TYPE "UDT_Service_StepRawDataMedium"
VERSION : 0.1
   STRUCT
      step { S7_SetPoint := 'False'} : Array[0..99] of "UDT_Service_StepMedium" := [([16#FFFFFFFF], [16#FFFFFFFF], [16#FFFFFFFF], [16#FFFFFFFF]), ([16#FFFFFFFF], [16#FFFFFFFF], [16#FFFFFFFF], [16#FFFFFFFF]), ([16#FFFFFFFF], [16#FFFFFFFF], [16#FFFFFFFF], [16#FFFFFFFF]), ([16#FFFFFFFF], [16#FFFFFFFF], [16#FFFFFFFF], [16#FFFFFFFF]), ([16#FFFFFFFF], [16#FFFFFFFF], [16#FFFFFFFF], [16#FFFFFFFF]), ([16#FFFFFFFF], [16#FFFFFFFF], [16#FFFFFFFF], [16#FFFFFFFF]), ([16#FFFFFFFF], [16#FFFFFFFF], [16#FFFFFFFF], [16#FFFFFFFF]), ([16#FFFFFFFF], [16#FFFFFFFF], [16#FFFFFFFF], [16#FFFFFFFF]), ([16#FFFFFFFF], [16#FFFFFFFF], [16#FFFFFFFF], [16#FFFFFFFF]), ([16#FFFFFFFF], [16#FFFFFFFF], [16#FFFFFFFF], [16#FFFFFFFF]), ([16#FFFFFFFF], [16#FFFFFFFF], [16#FFFFFFFF], [16#FFFFFFFF]), ([16#FFFFFFFF], [16#FFFFFFFF], [16#FFFFFFFF], [16#FFFFFFFF]), ([16#FFFFFFFF], [16#FFFFFFFF], [16#FFFFFFFF], [16#FFFFFFFF]), ([16#FFFFFFFF], [16#FFFFFFFF], [16#FFFFFFFF], [16#FFFFFFFF]), ([16#FFFFFFFF], [16#FFFFFFFF], [16#FFFFFFFF], [16#FFFFFFFF]), ([16#FFFFFFFF], [16#FFFFFFFF], [16#FFFFFFFF], [16#FFFFFFFF]), ([16#FFFFFFFF], [16#FFFFFFFF], [16#FFFFFFFF], [16#FFFFFFFF]), ([16#FFFFFFFF], [16#FFFFFFFF], [16#FFFFFFFF], [16#FFFFFFFF]), ([16#FFFFFFFF], [16#FFFFFFFF], [16#FFFFFFFF], [16#FFFFFFFF]), ([16#FFFFFFFF], [16#FFFFFFFF], [16#FFFFFFFF], [16#FFFFFFFF]), ([16#FFFFFFFF], [16#FFFFFFFF], [16#FFFFFFFF], [16#FFFFFFFF]), ([16#FFFFFFFF], [16#FFFFFFFF], [16#FFFFFFFF], [16#FFFFFFFF]), ([16#FFFFFFFF], [16#FFFFFFFF], [16#FFFFFFFF], [16#FFFFFFFF]), ([16#FFFFFFFF], [16#FFFFFFFF], [16#FFFFFFFF], [16#FFFFFFFF]), ([16#FFFFFFFF], [16#FFFFFFFF], [16#FFFFFFFF], [16#FFFFFFFF]), ([16#FFFFFFFF], [16#FFFFFFFF], [16#FFFFFFFF], [16#FFFFFFFF]), ([16#FFFFFFFF], [16#FFFFFFFF], [16#FFFFFFFF], [16#FFFFFFFF]), ([16#FFFFFFFF], [16#FFFFFFFF], [16#FFFFFFFF], [16#FFFFFFFF]), ([16#FFFFFFFF], [16#FFFFFFFF], [16#FFFFFFFF], [16#FFFFFFFF]), ([16#FFFFFFFF], [16#FFFFFFFF], [16#FFFFFFFF], [16#FFFFFFFF]), ([16#FFFFFFFF], [16#FFFFFFFF], [16#FFFFFFFF], [16#FFFFFFFF]), ([16#FFFFFFFF], [16#FFFFFFFF], [16#FFFFFFFF], [16#FFFFFFFF]), ([16#FFFFFFFF], [16#FFFFFFFF], [16#FFFFFFFF], [16#FFFFFFFF]), ([16#FFFFFFFF], [16#FFFFFFFF], [16#FFFFFFFF], [16#FFFFFFFF]), ([16#FFFFFFFF], [16#FFFFFFFF], [16#FFFFFFFF], [16#FFFFFFFF]), ([16#FFFFFFFF], [16#FFFFFFFF], [16#FFFFFFFF], [16#FFFFFFFF]), ([16#FFFFFFFF], [16#FFFFFFFF], [16#FFFFFFFF], [16#FFFFFFFF]), ([16#FFFFFFFF], [16#FFFFFFFF], [16#FFFFFFFF], [16#FFFFFFFF]), ([16#FFFFFFFF], [16#FFFFFFFF], [16#FFFFFFFF], [16#FFFFFFFF]), ([16#FFFFFFFF], [16#FFFFFFFF], [16#FFFFFFFF], [16#FFFFFFFF]), ([16#FFFFFFFF], [16#FFFFFFFF], [16#FFFFFFFF], [16#FFFFFFFF]), ([16#FFFFFFFF], [16#FFFFFFFF], [16#FFFFFFFF], [16#FFFFFFFF]), ([16#FFFFFFFF], [16#FFFFFFFF], [16#FFFFFFFF], [16#FFFFFFFF]), ([16#FFFFFFFF], [16#FFFFFFFF], [16#FFFFFFFF], [16#FFFFFFFF]), ([16#FFFFFFFF], [16#FFFFFFFF], [16#FFFFFFFF], [16#FFFFFFFF]), ([16#FFFFFFFF], [16#FFFFFFFF], [16#FFFFFFFF], [16#FFFFFFFF]), ([16#FFFFFFFF], [16#FFFFFFFF], [16#FFFFFFFF], [16#FFFFFFFF]), ([16#FFFFFFFF], [16#FFFFFFFF], [16#FFFFFFFF], [16#FFFFFFFF]), ([16#FFFFFFFF], [16#FFFFFFFF], [16#FFFFFFFF], [16#FFFFFFFF]), ([16#FFFFFFFF], [16#FFFFFFFF], [16#FFFFFFFF], [16#FFFFFFFF]), ([16#FFFFFFFF], [16#FFFFFFFF], [16#FFFFFFFF], [16#FFFFFFFF]), ([16#FFFFFFFF], [16#FFFFFFFF], [16#FFFFFFFF], [16#FFFFFFFF]), ([16#FFFFFFFF], [16#FFFFFFFF], [16#FFFFFFFF], [16#FFFFFFFF]), ([16#FFFFFFFF], [16#FFFFFFFF], [16#FFFFFFFF], [16#FFFFFFFF]), ([16#FFFFFFFF], [16#FFFFFFFF], [16#FFFFFFFF], [16#FFFFFFFF]), ([16#FFFFFFFF], [16#FFFFFFFF], [16#FFFFFFFF], [16#FFFFFFFF]), ([16#FFFFFFFF], [16#FFFFFFFF], [16#FFFFFFFF], [16#FFFFFFFF]), ([16#FFFFFFFF], [16#FFFFFFFF], [16#FFFFFFFF], [16#FFFFFFFF]), ([16#FFFFFFFF], [16#FFFFFFFF], [16#FFFFFFFF], [16#FFFFFFFF]), ([16#FFFFFFFF], [16#FFFFFFFF], [16#FFFFFFFF], [16#FFFFFFFF]), ([16#FFFFFFFF], [16#FFFFFFFF], [16#FFFFFFFF], [16#FFFFFFFF]), ([16#FFFFFFFF], [16#FFFFFFFF], [16#FFFFFFFF], [16#FFFFFFFF]), ([16#FFFFFFFF], [16#FFFFFFFF], [16#FFFFFFFF], [16#FFFFFFFF]), ([16#FFFFFFFF], [16#FFFFFFFF], [16#FFFFFFFF], [16#FFFFFFFF]), ([16#FFFFFFFF], [16#FFFFFFFF], [16#FFFFFFFF], [16#FFFFFFFF]), ([16#FFFFFFFF], [16#FFFFFFFF], [16#FFFFFFFF], [16#FFFFFFFF]), ([16#FFFFFFFF], [16#FFFFFFFF], [16#FFFFFFFF], [16#FFFFFFFF]), ([16#FFFFFFFF], [16#FFFFFFFF], [16#FFFFFFFF], [16#FFFFFFFF]), ([16#FFFFFFFF], [16#FFFFFFFF], [16#FFFFFFFF], [16#FFFFFFFF]), ([16#FFFFFFFF], [16#FFFFFFFF], [16#FFFFFFFF], [16#FFFFFFFF]), ([16#FFFFFFFF], [16#FFFFFFFF], [16#FFFFFFFF], [16#FFFFFFFF]), ([16#FFFFFFFF], [16#FFFFFFFF], [16#FFFFFFFF], [16#FFFFFFFF]), ([16#FFFFFFFF], [16#FFFFFFFF], [16#FFFFFFFF], [16#FFFFFFFF]), ([16#FFFFFFFF], [16#FFFFFFFF], [16#FFFFFFFF], [16#FFFFFFFF]), ([16#FFFFFFFF], [16#FFFFFFFF], [16#FFFFFFFF], [16#FFFFFFFF]), ([16#FFFFFFFF], [16#FFFFFFFF], [16#FFFFFFFF], [16#FFFFFFFF]), ([16#FFFFFFFF], [16#FFFFFFFF], [16#FFFFFFFF], [16#FFFFFFFF]), ([16#FFFFFFFF], [16#FFFFFFFF], [16#FFFFFFFF], [16#FFFFFFFF]), ([16#FFFFFFFF], [16#FFFFFFFF], [16#FFFFFFFF], [16#FFFFFFFF]), ([16#FFFFFFFF], [16#FFFFFFFF], [16#FFFFFFFF], [16#FFFFFFFF]), ([16#FFFFFFFF], [16#FFFFFFFF], [16#FFFFFFFF], [16#FFFFFFFF]), ([16#FFFFFFFF], [16#FFFFFFFF], [16#FFFFFFFF], [16#FFFFFFFF]), ([16#FFFFFFFF], [16#FFFFFFFF], [16#FFFFFFFF], [16#FFFFFFFF]), ([16#FFFFFFFF], [16#FFFFFFFF], [16#FFFFFFFF], [16#FFFFFFFF]), ([16#FFFFFFFF], [16#FFFFFFFF], [16#FFFFFFFF], [16#FFFFFFFF]), ([16#FFFFFFFF], [16#FFFFFFFF], [16#FFFFFFFF], [16#FFFFFFFF]), ([16#FFFFFFFF], [16#FFFFFFFF], [16#FFFFFFFF], [16#FFFFFFFF]), ([16#FFFFFFFF], [16#FFFFFFFF], [16#FFFFFFFF], [16#FFFFFFFF]), ([16#FFFFFFFF], [16#FFFFFFFF], [16#FFFFFFFF], [16#FFFFFFFF]), ([16#FFFFFFFF], [16#FFFFFFFF], [16#FFFFFFFF], [16#FFFFFFFF]), ([16#FFFFFFFF], [16#FFFFFFFF], [16#FFFFFFFF], [16#FFFFFFFF]), ([16#FFFFFFFF], [16#FFFFFFFF], [16#FFFFFFFF], [16#FFFFFFFF]), ([16#FFFFFFFF], [16#FFFFFFFF], [16#FFFFFFFF], [16#FFFFFFFF]), ([16#FFFFFFFF], [16#FFFFFFFF], [16#FFFFFFFF], [16#FFFFFFFF]), ([16#FFFFFFFF], [16#FFFFFFFF], [16#FFFFFFFF], [16#FFFFFFFF]), ([16#FFFFFFFF], [16#FFFFFFFF], [16#FFFFFFFF], [16#FFFFFFFF]), ([16#FFFFFFFF], [16#FFFFFFFF], [16#FFFFFFFF], [16#FFFFFFFF]), ([16#FFFFFFFF], [16#FFFFFFFF], [16#FFFFFFFF], [16#FFFFFFFF]), ([16#FFFFFFFF], [16#FFFFFFFF], [16#FFFFFFFF], [16#FFFFFFFF]), ([16#FFFFFFFF], [16#FFFFFFFF], [16#FFFFFFFF], [16#FFFFFFFF])];
      parameterDefinition { S7_SetPoint := 'False'} : Array[0..31] of "UDT_Service_ParameterDefinition";
   END_STRUCT;

END_TYPE

